FUNCTION F_ConvertSetPosResiduals : DINT
(*
Convert technical units to inc

*)
VAR_INPUT

	(* Enummerations *)
	
	(* Variables *)
	lrPos								:LREAL;

	(* References *)

	(* Interfaces *)
	pAxis								:POINTER TO ST_AXIS_REF_V2;

	(* Instances *)

END_VAR
VAR
END_VAR


IF pAxis^.stScaling.etScalingMethod = ET_ScalingMethod_eSMRotary
THEN

	F_ConvertSetPosResiduals := LREAL_TO_DINT(lrPos);

ELSIF pAxis^.stScaling.etScalingMethod = ET_ScalingMethod_eSMLinear
THEN

	F_ConvertSetPosResiduals := LREAL_TO_DINT((lrPos + pAxis^.stPosition.lrOffsetPos) * pAxis^.stScaling.lrScaleFactor);

END_IF

IF pAxis^.stScaling.dwModuloValue > 0
THEN
	F_ConvertSetPosResiduals := DWORD_TO_DINT(DINT_TO_DWORD(F_ConvertSetPosResiduals) MOD pAxis^.stScaling.dwModuloValue);
END_IF

END_FUNCTION

(* stored: Version 1.1.0.1, ProductVersion 3.1.4024.15
   POU F_ConvertSetPosResiduals: Id {a3666087-d9f1-41aa-9f0a-e289135149aa}, SpecialFunc None *)
